(* PLC project Vn_ton_in_box, Beckhoff Automation GmbH TwinCAT PLC Control 3.5.13.21 *)
(* stored: creationDateTime 1970-01-01T00:00:00 *)

PROGRAM Vn_ton_in_box

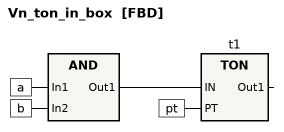
(* FBD diagram, written out as Structured Text *)
t1(IN := a AND b, PT := pt);
END_PROGRAM
